(* IEC 61131-3 sources: factory_in_a_box/firmware_factory_control_unit/web_packages/plc/src/corpus, 26 files *)

(* ---- fb_user.st ---- *)
(* @cycles 20 *)
FUNCTION_BLOCK FB_PID
VAR_INPUT sp : REAL; pv : REAL; kp : REAL := 1.0; ki : REAL := 0.1; END_VAR
VAR_OUTPUT y : REAL; END_VAR
VAR i : REAL; END_VAR
i := LIMIT(-50.0, i + ki * (sp - pv), 50.0);
y := kp * (sp - pv) + i;
END_FUNCTION_BLOCK
FUNCTION_BLOCK FB_PLANT
VAR_INPUT u : REAL; END_VAR
VAR_OUTPUT x : REAL; END_VAR
x := x + 0.2 * (u - x);
END_FUNCTION_BLOCK
PROGRAM PLC_PRG
VAR c : FB_PID; p : FB_PLANT; ctl : ARRAY[0..1] OF FB_PID; y2 : REAL; END_VAR
c(sp := 10.0, pv := p.x);
p(u := c.y);
ctl[1](sp := 5.0, pv := y2, kp := 0.5, y => y2);
END_PROGRAM

(* ---- nested_fb_std.st ---- *)
(* @cycles 30 *)
(* @dt 25 *)
FUNCTION_BLOCK FB_BLINK
VAR_INPUT en : BOOL; period : TIME := T#100ms; END_VAR
VAR_OUTPUT q : BOOL; toggles : INT; END_VAR
VAR t : TON; END_VAR
t(IN := en AND NOT t.Q, PT := period / 2);
IF t.Q THEN q := NOT q; toggles := toggles + 1; END_IF;
END_FUNCTION_BLOCK
PROGRAM PLC_PRG
VAR b1 : FB_BLINK; b2 : FB_BLINK; both : INT; END_VAR
b1(en := TRUE);
b2(en := TRUE, period := T#250ms);
IF b1.q AND b2.q THEN both := both + 1; END_IF;
END_PROGRAM

(* ---- array_trap.st ---- *)
(* @cycles 10 *)
PROGRAM PLC_PRG
VAR a : ARRAY[2..6] OF DINT; i : INT := 2; END_VAR
a[i] := i * 10;
i := i + 1;
END_PROGRAM

(* ---- bits.st ---- *)
(* @cycles 20 *)
PROGRAM PLC_PRG
VAR b : BYTE := 16#81; w : WORD := 16#8001; d : DWORD := 16#80000001; l : LWORD := 16#8000000000000001;
    sb : BYTE; sw : WORD; rd : DWORD; rl : LWORD; x : DWORD; n : INT; m : BOOL; END_VAR
sb := SHL(b, n); sw := SHR(w, n); rd := ROL(d, n); rl := ROR(l, n);
x := (d AND 16#FF00FF00) OR (DWORD#16#00F0F0F0 XOR rd);
b := ROL(b, 3); w := NOT w; l := l XOR SHL(l, 1);
m := (b AND 16#01) = 16#01;
n := n + 1;
END_PROGRAM

(* ---- budget_trap.st ---- *)
(* @cycles 3 *)
(* @budget 5000 *)
PROGRAM PLC_PRG
VAR n : DINT; END_VAR
WHILE n >= 0 DO n := n + 1; END_WHILE;
END_PROGRAM

(* ---- case_enum.st ---- *)
(* @cycles 12 *)
TYPE E_State : (Idle, Fill, Heat := 10, Drain, Done); END_TYPE
PROGRAM PLC_PRG
VAR st : E_State; t : INT; n : INT; hist : ARRAY[0..11] OF E_State; c : INT; END_VAR
CASE st OF
  Idle: st := Fill;
  Fill: t := t + 1; IF t >= 3 THEN st := Heat; t := 0; END_IF;
  Heat, Drain: t := t + 2; IF t > 3 THEN st := SEL(st = Heat, Done, Drain); t := 0; END_IF;
ELSE
  st := Idle;
END_CASE;
CASE n OF
  0..2: c := 1;
  3, 5, 7: c := 2;
  -5..-1: c := 3;
ELSE c := 4;
END_CASE;
hist[n] := st;
n := n + 1;
END_PROGRAM

(* ---- conv_double_rounding.st ---- *)
(* @cycles 2 *)
PROGRAM PLC_PRG
VAR v : LINT := 1152921573326323713; f : REAL; g : REAL; uv : ULINT := 18446744073709551615; h : REAL; hl : LREAL; END_VAR
(* 2^60 + 2^36 + 1: rounded once to REAL gives 2^60 + 2^37 *)
f := LINT_TO_REAL(v); g := LINT_TO_REAL(-v); h := ULINT_TO_REAL(uv); hl := ULINT_TO_LREAL(uv);
v := v + 1;
END_PROGRAM

(* ---- conv_trap.st ---- *)
(* @cycles 10 *)
PROGRAM PLC_PRG
VAR d : DINT := 32760; i : INT; END_VAR
i := DINT_TO_INT(d);
d := d + 1;
END_PROGRAM

(* ---- conversions.st ---- *)
(* @cycles 25 *)
PROGRAM PLC_PRG
VAR r : REAL := -12.5; lr : LREAL := 1.0E15; i : INT; d : DINT; l : LINT; ul : ULINT; t : DINT;
    rr : REAL; lrr : LREAL; b : BOOL; w : WORD; dw : DWORD; si : SINT; k : DINT := -3; END_VAR
i := REAL_TO_INT(r); d := TRUNC(r); l := LREAL_TO_LINT(lr); t := REAL_TO_DINT(r * 1000.0);
rr := DINT_TO_REAL(k * 33333); lrr := LINT_TO_LREAL(l * 3);
b := INT_TO_BOOL(i); w := INT_TO_WORD(i); dw := WORD_TO_DWORD(w); si := WORD_TO_SINT(w);
ul := LINT_TO_ULINT(ABS(l));
r := r + 1.0; lr := lr * 3.0; k := k * 7;
END_PROGRAM

(* ---- counter.st ---- *)
(* @cycles 10 *)
(* @expect PLC_PRG.n = 10 *)
PROGRAM PLC_PRG
VAR n : DINT; END_VAR
n := n + 1;
END_PROGRAM

(* ---- counters_edges.st ---- *)
(* @cycles 40 *)
PROGRAM PLC_PRG
VAR clk : BOOL; n : INT; up : CTU; dn : CTD; ud : CTUD; r : R_TRIG; f : F_TRIG; s : SR; rs : RS; edges : INT; END_VAR
clk := (n MOD 3) = 0;
r(CLK := clk); f(CLK := clk);
IF r.Q OR f.Q THEN edges := edges + 1; END_IF;
up(CU := clk, R := n = 25, PV := 5);
dn(CD := clk, LD := n = 0, PV := 4);
ud(CU := clk, CD := NOT clk AND (n MOD 5 = 0), R := FALSE, LD := FALSE, PV := 3);
s(S1 := n = 10, R := n = 20); rs(S := n = 12, R1 := n = 15);
n := n + 1;
END_PROGRAM

(* ---- div_zero_trap.st ---- *)
(* @cycles 10 *)
PROGRAM PLC_PRG
VAR a : DINT := 100; b : DINT := 4; c : DINT; END_VAR
c := a / b;
b := b - 1;
END_PROGRAM

(* ---- functions.st ---- *)
(* @cycles 6 *)
FUNCTION CLAMP_ADD : INT
VAR_INPUT a : INT; b : INT; lo : INT := -100; hi : INT := 100; END_VAR
CLAMP_ADD := LIMIT(lo, a + b, hi);
END_FUNCTION
FUNCTION POLY : LREAL
VAR_INPUT x : LREAL; END_VAR
VAR c : ARRAY[0..3] OF LREAL := [1.0, -2.0, 0.5, 0.25]; i : INT; END_VAR
FOR i := 3 TO 0 BY -1 DO POLY := POLY * x + c[i]; END_FOR;
END_FUNCTION
FUNCTION SWAP2 : BOOL
VAR_IN_OUT a : DINT; b : DINT; END_VAR
VAR t : DINT; END_VAR
t := a; a := b; b := t; SWAP2 := a > b;
END_FUNCTION
FUNCTION DEPTH : DINT
VAR_INPUT n : DINT; END_VAR
DEPTH := n + POLY_INT(n);
END_FUNCTION
FUNCTION POLY_INT : DINT
VAR_INPUT n : DINT; END_VAR
POLY_INT := LREAL_TO_DINT(POLY(DINT_TO_LREAL(n)));
END_FUNCTION
PROGRAM PLC_PRG
VAR s : INT; p : LREAL; x : DINT := 5; y : DINT := 9; g : BOOL; d : DINT; END_VAR
s := CLAMP_ADD(a := s, b := 37); s := CLAMP_ADD(a := s, b := -5, hi := 120);
p := POLY(INT_TO_LREAL(s) / 10.0);
g := SWAP2(x, y);
d := DEPTH(x);
END_PROGRAM

(* ---- globals.st ---- *)
(* @cycles 7 *)
VAR_GLOBAL
  g_count : UDINT := 1000;
  g_tab : ARRAY[0..4] OF INT := [5, 4, 3, 2(9)];
END_VAR
VAR_GLOBAL CONSTANT
  K : INT := 4;
END_VAR
PROGRAM PLC_PRG
VAR i : INT; mx : INT; mn : INT; mu : INT; n : INT; END_VAR
g_count := g_count * 3;
FOR i := 0 TO K DO g_tab[i] := g_tab[i] + i; END_FOR;
mx := MAX(g_tab[0], g_tab[1], g_tab[2], g_tab[3], g_tab[4]);
mn := MIN(g_tab[0], g_tab[4]);
mu := MUX(n, 11, 22, 33, 44, 55, 66, 77);
n := n + 1;
END_PROGRAM

(* ---- int_compare.st ---- *)
(* @cycles 40 *)
PROGRAM PLC_PRG
VAR i : INT := -20; u : UDINT := 4294967270; l : LINT := -5; ul : ULINT := 18446744073709551590;
    c1 : BOOL; c2 : BOOL; c3 : BOOL; c4 : BOOL; c5 : BOOL; c6 : BOOL; n : DINT; END_VAR
c1 := i < 0; c2 := u > 4294967282; c3 := l <= -3; c4 := ul >= 18446744073709551602; c5 := i <> 0; c6 := (i = 0) OR (u = 0);
IF c1 THEN n := n + 1; END_IF;
IF c2 AND c4 THEN n := n + 100; END_IF;
i := i + 1; u := u + 1; l := l + 1; ul := ul + 1;
END_PROGRAM

(* ---- int_divmod.st ---- *)
(* @cycles 30 *)
PROGRAM PLC_PRG
VAR a : DINT := -1000; b : DINT := 7; q : DINT; r : DINT; ua : UDINT := 4000000000; uq : UDINT; ur : UDINT;
    la : LINT := -9000000000000; lq : LINT; lr : LINT; ula : ULINT := 18000000000000000000; ulq : ULINT; si : SINT := -128; sq : SINT; END_VAR
q := a / b; r := a MOD b; uq := ua / DINT_TO_UDINT(b); ur := ua MOD 13;
lq := la / 13; lr := la MOD 13; ulq := ula / 3;
sq := si / -1;
a := a + 77; b := b + 1; ua := ua - 12345; la := la * 3;
END_PROGRAM

(* ---- int_wrap.st ---- *)
(* @cycles 300 *)
(* @expect PLC_PRG.s = 44 *)
(* @expect PLC_PRG.u = 44 *)
PROGRAM PLC_PRG
VAR s : SINT; u : USINT; i : INT := 32700; w : UINT := 65500; d : DINT := 2147483600; l : LINT := 9223372036854775800; ul : ULINT := 18446744073709551600; END_VAR
s := s + 1; u := u + 1; i := i + 1; w := w + 1; d := d + 1; l := l + 1; ul := ul + 1;
END_PROGRAM

(* ---- loops.st ---- *)
(* @cycles 5 *)
PROGRAM PLC_PRG
VAR i : INT; j : INT; s : DINT; st : INT := -2; k : INT; fib : ARRAY[0..20] OF DINT; END_VAR
FOR i := 1 TO 10 DO FOR j := i TO 10 BY 3 DO s := s + i * j; END_FOR; END_FOR;
FOR i := 9 TO 0 BY st DO s := s - i; END_FOR;
fib[0] := 0; fib[1] := 1;
FOR i := 2 TO 20 DO fib[i] := fib[i - 1] + fib[i - 2]; END_FOR;
k := 0;
REPEAT k := k + 1; IF k = 3 THEN CONTINUE; END_IF; s := s + k; UNTIL k > 6 END_REPEAT;
WHILE TRUE DO s := s + 1; IF s MOD 7 = 0 THEN EXIT; END_IF; END_WHILE;
END_PROGRAM

(* ---- lreal_math.st ---- *)
(* @cycles 20 *)
PROGRAM PLC_PRG
VAR x : LREAL := 2.0; s : LREAL; e : LREAL; a : LREAL; r : REAL := 2.0; sr : REAL; k : INT := -7; ak : INT; END_VAR
s := SQRT(x); sr := SQRT(r); x := x * 1.5 + s;
e := s * s;
a := ABS(-x); ak := ABS(k); k := k + 1;
r := r * 1.25;
END_PROGRAM

(* ---- multi_program.st ---- *)
(* @cycles 6 *)
(* @programs PLC_PRG P2 *)
VAR_GLOBAL shared : DINT; END_VAR
PROGRAM PLC_PRG
VAR n : DINT; END_VAR
n := n + 1; shared := shared * 2 + n;
END_PROGRAM
PROGRAM P2
VAR last : DINT; END_VAR
last := shared; shared := shared - 1;
END_PROGRAM

(* ---- real_arith.st ---- *)
(* @cycles 50 *)
PROGRAM PLC_PRG
VAR x : REAL := 0.1; y : REAL := 3.0; s : REAL; p : REAL := 1.0; q : REAL; big : REAL := 1.0E30; tiny : REAL := 1.0E-30;
    lx : LREAL := 0.1; ls : LREAL; lp : LREAL := 1.0; c : BOOL; END_VAR
s := s + x; p := p * 1.1; q := s / y; big := big * 7.0; tiny := tiny / 3.0;
ls := ls + lx; lp := lp * 1.0000001;
c := s > q;
x := x + 0.07;
END_PROGRAM

(* ---- real_special.st ---- *)
(* @cycles 3 *)
PROGRAM PLC_PRG
VAR a : REAL := -1.0; n1 : REAL; n2 : LREAL; inf : REAL := 3.0E38; i2 : REAL; ninf : REAL; z : REAL; c1 : BOOL; c2 : BOOL; c3 : BOOL; ab : REAL; END_VAR
n1 := SQRT(a); n2 := SQRT(REAL_TO_LREAL(a));
i2 := inf * 10.0; ninf := -i2; z := i2 + ninf;
c1 := n1 = n1; c2 := n1 <> n1; c3 := z < 0.0;
ab := ABS(ninf);
END_PROGRAM

(* ---- structs_arrays.st ---- *)
(* @cycles 8 *)
TYPE
  S_Point : STRUCT x : INT := 1; y : INT := -1; END_STRUCT;
  S_Path : STRUCT p : ARRAY[0..3] OF S_Point; len : USINT := 4; name : DWORD := 16#CAFE; END_STRUCT;
END_TYPE
PROGRAM PLC_PRG
VAR a : S_Path; b : S_Path; m : ARRAY[1..3, 1..4] OF LREAL; i : INT := 1; j : INT := 1; k : INT; tot : LREAL; END_VAR
a.p[k].x := a.p[k].x + k; a.p[3 - k].y := a.p[k].x * 2;
b := a;
m[i, j] := INT_TO_LREAL(a.p[k].x) / 3.0;
tot := tot + m[i, j];
j := j + 1; IF j > 4 THEN j := 1; i := i + 1; END_IF;
k := (k + 1) MOD 4;
END_PROGRAM

(* ---- subrange_trap.st ---- *)
(* @cycles 20 *)
TYPE T_Pct : INT (0..100); END_TYPE
PROGRAM PLC_PRG
VAR p : T_Pct := 40; END_VAR
p := p + 7;
END_PROGRAM

(* ---- time_ops.st ---- *)
(* @cycles 10 *)
(* @dt 37 *)
PROGRAM PLC_PRG
VAR t : TIME := T#1h2m3s4ms; u : TIME; n : DINT := 3; d : DINT; neg : TIME := T#-1500ms; c : BOOL; END_VAR
u := t * n - T#1d / 4 + neg;
d := TIME_TO_DINT(u);
c := u > T#0ms;
t := t / 2;
END_PROGRAM

(* ---- timers.st ---- *)
(* @cycles 60 *)
(* @dt 10 *)
(* @set 5 PLC_PRG.in := 1 *)
(* @set 30 PLC_PRG.in := 0 *)
(* @set 33 PLC_PRG.in := 1 *)
(* @set 35 PLC_PRG.in := 0 *)
(* @expect PLC_PRG.ton_q_cycles = 16 *)
PROGRAM PLC_PRG
VAR in : BOOL; t1 : TON; t2 : TOF; t3 : TP; ton_q_cycles : INT; tof_q : INT; tp_q : INT; END_VAR
t1(IN := in, PT := T#90ms); t2(IN := in, PT := T#40ms); t3(IN := in, PT := T#70ms);
IF t1.Q THEN ton_q_cycles := ton_q_cycles + 1; END_IF;
IF t2.Q THEN tof_q := tof_q + 1; END_IF;
IF t3.Q THEN tp_q := tp_q + 1; END_IF;
END_PROGRAM
